Fanuc KAREL source: KX00031.KL

PROGRAM KX00031
%NOLOCKGROUP
%DEFGROUP = 1
VAR
  I: INTEGER
  J: INTEGER
  B: BOOLEAN
  F: FILE
  S: STRING[80]
  P: XYZWPR
BEGIN
  I = 1
END KX00031
